// TIA Portal V20 export
Screen "190FX2RhSliderLayout"  1276x673
  ScreenItem "Line_Header_X0_Y64" at 0,64 size 1276x0  Type=HmiLine
  ScreenItem "permanentareaborderrectangle" at 0,0 size 0x0  Type=HmiRectangle
  ScreenItem "Button_Back" at 2,2 size 90x60  Type=HmiButton
  ScreenItem "Move_Legend" at 1182,2 size 90x60  Type=HmiButton
  ScreenItem "Fusszeile_Button_ManualOPMode1_2" at 279,2 size 90x60  Type=HmiButton
  ScreenItem "文本域_3" at 1109,71 size 139x22  Type=HmiTextBox
  ScreenItem "文本域_1" at 1101,160 size 156x23  Type=HmiTextBox
  ScreenItem "文本域_2" at 1111,246 size 135x23  Type=HmiTextBox
  ScreenItem "文本域_22" at 1129,384 size 104x23  Type=HmiTextBox
  ScreenItem "Fusszeile_Button_ManualOPMode1_1" at 95,2 size 90x60  Type=HmiButton
  ScreenItem "Button_Back_1" at 1180,606 size 90x60  Type=HmiButton
  ScreenItem "Fusszeile_Button_ManualOPMode1_3" at 187,2 size 90x60  Type=HmiButton
  ScreenItem "Fusszeile_Button_ManualOPMode1_4" at 997,2 size 90x60  Type=HmiButton
  ScreenItem "Fusszeile_Button_ManualOPMode1_5" at 902,1 size 90x60  Type=HmiButton
  ScreenItem "文本域_14" at 936,-172 size 140x40  Type=HmiTextBox
  ScreenItem "Graphic view_1" at 226,212 size 651x296  Type=HmiGraphicView
  ScreenItem "文本域_5" at -1,82 size 120x40  Type=HmiTextBox
  ScreenItem "文本域_27" at -1,126 size 120x40  Type=HmiTextBox
  ScreenItem "LSicar_Valve8Pos_LeftHomeRightWork_WithPB_5" at 1099,95 size 160x53  Type=HmiFaceplateContainer
  ScreenItem "LSicar_Valve8Pos_LeftHomeRightWork_WithPB_1" at 1099,183 size 160x53  Type=HmiFaceplateContainer
  ScreenItem "面板容器_22" at 1066,417 size 96x32  Type=HmiFaceplateContainer
  ScreenItem "面板容器_23" at 1176,417 size 96x32  Type=HmiFaceplateContainer
  ScreenItem "LSicar_Valve8Pos_LeftHomeRightWork_WithPB_2" at 1099,271 size 160x53  Type=HmiFaceplateContainer
  ScreenItem "文本域_21" at 256,107 size 140x40  Type=HmiTextBox
  ScreenItem "Line_4" at 356,173 size 115x131  Type=HmiLine
  ScreenItem "文本域_12" at 532,109 size 100x40  Type=HmiTextBox
  ScreenItem "Line_1" at 487,190 size 78x207  Type=HmiLine
  ScreenItem "文本域_6" at 55,309 size 140x40  Type=HmiTextBox
  ScreenItem "面板容器_1" at 59,357 size 144x51  Type=HmiFaceplateContainer
  ScreenItem "Line_2" at 200,341 size 197x112  Type=HmiLine
  ScreenItem "文本域_7" at 924,309 size 100x40  Type=HmiTextBox
  ScreenItem "Faceplate container_1" at 944,357 size 59x45  Type=HmiFaceplateContainer
  ScreenItem "Line_3" at 844,334 size 78x43  Type=HmiLine
  ScreenItem "文本域_8" at 815,557 size 100x40  Type=HmiTextBox
  ScreenItem "Faceplate container_2" at 835,597 size 59x45  Type=HmiFaceplateContainer
  ScreenItem "Line_5" at 573,434 size 239x144  Type=HmiLine
  ScreenItem "文本域_9" at 577,557 size 100x40  Type=HmiTextBox
  ScreenItem "Faceplate container_3" at 597,597 size 59x45  Type=HmiFaceplateContainer
  ScreenItem "Line_6" at 530,502 size 82x52  Type=HmiLine
  ScreenItem "文本域_10" at 359,557 size 100x40  Type=HmiTextBox
  ScreenItem "Faceplate container_4" at 379,597 size 59x45  Type=HmiFaceplateContainer
  ScreenItem "Line_7" at 426,473 size 62x82  Type=HmiLine
  ScreenItem "Title_ScreenOverview_X390_Y2_1" at 384,5 size 510x57  Type=HmiTextBox
  ScreenItem "面板容器_8" at 258,148 size 144x51  Type=HmiFaceplateContainer
  ScreenItem "Button_Back_2" at 1077,606 size 90x60  Type=HmiButton
  ScreenItem "Faceplate container_6" at 552,149 size 59x45  Type=HmiFaceplateContainer
  ScreenItem "面板容器_2" at 1090,4 size 88x58  Type=HmiFaceplateContainer
  ScreenItem "OPMode1_Blocked" at 1164,6 size 14x14  Type=HmiGraphicView
  ScreenItem "OPMode4_Foreground_Blocked" at 1089,2 size 88x58  Type=HmiGraphicView
